(*
SPDX-FileCopyrightText: © 2026 Oleksandr Tiutyk <trofimich@gmail.com>
SPDX-License-Identifier: MIT
License: https://opensource.org/license/mit
*)

(*!
<summary>Runs one single-cycle test directly, without a group.</summary>
<description>
Map this program to one cyclic PLC task or call its Execute method once per cycle from that task.
The concrete runner owns the tests; the program owns the reporter and performs task
cleanup at the end of every scan. Inspect _Runner.IsFinished, AllPassed and counts, then _Report.IsReady.
For independent task execution, assign SingleCycleTestExample and MultiCycleTestExample to different tasks.
They share no instances or mutable buffers. Do not assign the same program instance to multiple tasks.
</description>
*)

{attribute 'no_explicit_call' := 'do not call this function block directly'}
PROGRAM SingleCycleTestExample
VAR
	{attribute 'hide'}
	_ClassName : STRING := __POUNAME();

	_Runner : AdditionTestRunner;
	_Report : TOF_Testing.JUnitXmlReporter;
	_Configured : BOOL;
END_VAR

Execute();

//! <summary>Borrows the concrete program name for its lifetime; callers must not modify it.</summary>
{attribute 'monitoring' := 'call'}
PROPERTY ClassName : REFERENCE TO STRING
GET
ClassName REF= _ClassName;
END_GET
END_PROPERTY

(*!
<summary>Advances this example and performs standalone task-boundary memory cleanup.</summary>
<description>
Call once per cycle from the owning task, either through this method or by mapping this PROGRAM to that task.
Do not drive both entry paths or share the instance between tasks. Use as the standalone example in its task;
hosts with additional transient-exception consumers must provide a shared boundary instead.
</description>
*)
METHOD Execute
IF NOT _Configured THEN
	_Runner.Reporter := _Report;
	_Configured := TRUE;
END_IF

_Runner.Execute(cleanupTaskMemory := TRUE);
END_METHOD

(*!
<summary>Provides the library namespace used in diagnostics.</summary>
<description>
Borrowed read-only reference to the compiler-initialized library namespace; no ownership transfer.
</description>
*)
{attribute 'monitoring' := 'call'}
PROPERTY NamespaceName : REFERENCE TO STRING
GET
NamespaceName REF= CurrentNamespace.Name;
END_GET
END_PROPERTY

END_PROGRAM

(* stored: Version 1.1.0.1
   POU SingleCycleTestExample: Id {36ea0b94-7266-4356-99dc-c1a204131fc8}, SpecialFunc None
   Property ClassName: Id {2d513973-13f2-4b02-a22d-8638e933b171}
   Get Get: Id {a3ba236b-03ef-49ea-ac08-79f1f908b24f}
   Method Execute: Id {871dd4f9-9f87-4f78-b8b9-38f0871de851}
   Property NamespaceName: Id {44d17294-f805-4713-8be6-69fc055ac5d1}
   Get Get: Id {c1494ddc-d7f7-44d3-9335-22322bbbed3b} *)
